// SIMATIC S7-200 project (STEP 7-Micro/WIN), CPU 224XP CN REL 02.01

SYMBOL_TABLE 用户定义1
Codificador_A    I0.0
Codificador_B    I0.1
Codificador_Z    I0.2
S_foto_banda     I0.3
S_Fibra_optica   I0.4
S_de_metal       I0.5
Piston_1         I0.7
Piston_2         I1.0
Piston_3         I1.1
Boton_rojo       I1.2
Boton_verde      I1.3
Boton_emergencia I1.4
Switch           I1.5
Listo            M0.0
Comienzo         M0.1
Piezas_metalicas M1.0
Centro           M1.1
Centro_metalico  M1.2
Centro_plastico  M1.3
Otro             M1.4
Variador_Start_Stop Q0.0
Solenoide_1      Q0.4
Solenoide_2      Q0.5
Solenoide_3      Q0.6
Foco_amarillo    Q0.7
Foco_verde       Q1.0
Foco_rojo        Q1.1
Solicitar_alimentacion V1000.4
Permitir_clasificacion V1000.7
Detener_la_produccion V1001.0
Paquete_despejado V1001.2
Red_normal       V1010.0
Funcionamiento_continuo V1010.1
Detener_completado V1010.2
Producieron_varios VB1011
Frec_inversor    VW1002
END_SYMBOL_TABLE

ORGANIZATION_BLOCK Principal:OB1
TITLE=
BEGIN
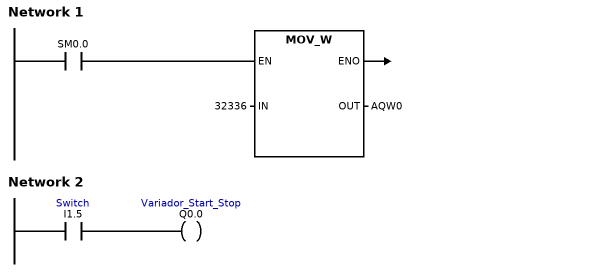
Network 1
LD     SM0.0
MOVW   32336, AQW0
Network 2
LD     Switch:I1.5
=      Variador_Start_Stop:Q0.0
END_ORGANIZATION_BLOCK

SUBROUTINE_BLOCK HSC_INIT:SBR1
TITLE=
BEGIN
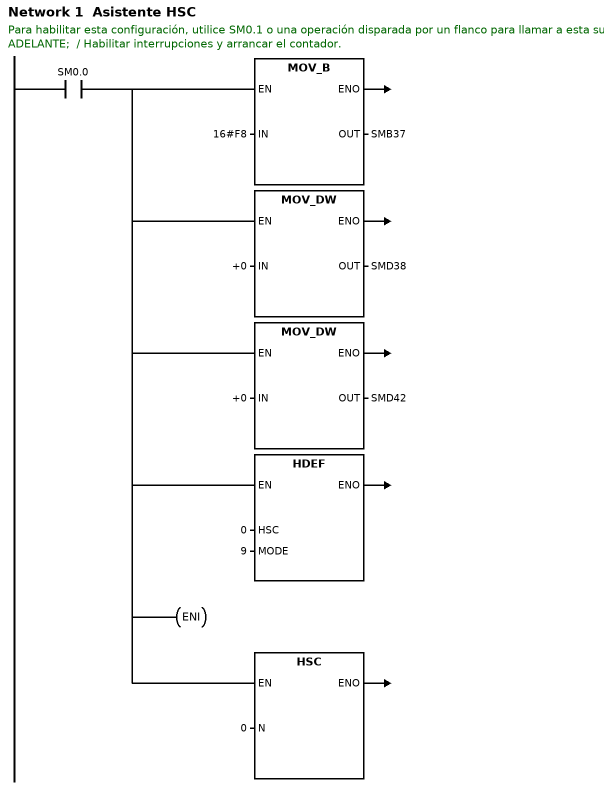
Network 1 // Asistente HSC 
// Para habilitar esta configuración, utilice SM0.1 o una operación disparada por un flanco para llamar a esta subrutina una vez desde el programa PRINCIPAL. 
// Configurar HC1 para modo 9; contar ADELANTE; 
// Habilitar interrupciones y arrancar el contador.
//设置控制位：增计数；4X 速率；已使能；
//装载 CV
//装载 PV
LD     SM0.0
MOVB   16#F8, SMB37
MOVD   +0, SMD38
MOVD   +0, SMD42
HDEF   0, 9
ENI
HSC    0
END_SUBROUTINE_BLOCK
